Fanuc KAREL source: KO00022.KL

PROGRAM KO00022
%NOLOCKGROUP
VAR
  P1: XYZWPREXT
  P2: XYZWPREXT
  P3: XYZWPREXT
  P4: XYZWPREXT
  OUT: XYZWPR
BEGIN
  OUT = FRAME(P1, P2, P3, P4)
END KO00022
